PROGRAM MAIN
VAR
    fbMessage1 : FB_MY_EVENT_MESSAGE;
    fbMessage2 : FB_MY_EVENT_MESSAGE;

    nError1 : UDINT := 0;
    nError2 : UDINT := 0;

    sError1 : T_MaxString := 'Testfehler Wechselrichter';
    sError2 : T_MaxString := 'Testfehler Speicher';

    nNow : Tc2_EtherCAT.T_DCTIME64;
	
	fbTiming1 : FB_MyTimingSample;
	fbTiming2 : FB_MyTimingSample;
	
	fbBase1 : FB_Base;
    fbBase2 : FB_Base;
    fbBase3 : FB_Base;
	
	nErrorFromRegister : UDINT;
END_VAR

// Aktuelle DC-Zeit.
// Der Meldungsbaustein speichert sie beim Erkennen eines Fehlers.
nNow := Tc2_EtherCAT.F_GetCurDcTickTime64();

fbMessage1(
    sSourcename := 'Wechselrichter',
    eLevel     := Tc3_EventLogger.TcEventSeverity.Error,
    nEventCode := TC_EVENTS.EC_Uebungen.ExternalError.nEventId,
    nError     := nError1,
    sError     := sError1,
    nTimeStamp := nNow
);

fbMessage2(
    sSourcename := 'Speicher',
    eLevel     := Tc3_EventLogger.TcEventSeverity.Warning,
    nEventCode := TC_EVENTS.EC_Uebungen.ExternalError.nEventId,
    nError     := nError2,
    sError     := sError2,
    nTimeStamp := nNow
);

IF GVL.Register.arrRegister[1] <> 0 THEN
    nErrorFromRegister := GVL.Register.arrRegister[1].Error;
END_IF

END_PROGRAM

(* stored: Version 1.1.0.1, ProductVersion 3.1.4024.16
   POU MAIN: Id {dcf70471-313e-4d4f-97bc-df7c8323bc4b}, SpecialFunc None *)
